(* IEC 61131-3 sources: JingjiangMoonbox/Application/Application/数据类型/通讯协议/月影/副主站通讯协议#1, 7 files *)

(* ---- StParam_Mailbox_Dep.st ---- *)
(*@CES
Name=StParam_Mailbox_Dep
Type=Gvl
TypeGuid=2db5746d-d284-4425-9f7f-2663a34b0ebc
Guid=8959721b-aa70-4a50-8488-8b5c585a49ff
HasDeclaration=True
HasImplementation=False
*)
{DECLARATION}
{attribute 'pack_mode' := '1'}
TYPE StParam_Mailbox_Dep :
STRUCT
	dwSemaphore								:DWORD;(*通讯旗语						*)

	iGirth_Uw_A								: INT; (*放A周长*)
	iGirth_Uw_B								: INT; (*放B周长*)
	iGirth_Pu								: INT;(*版周长*)
	iVelocity_Tar							: INT;(*目标速度*)
	iAI_mid_Uw								: INT;(*放料中位*)
	iAI_mid_If								: INT;(*放牵中位*)
	byDir_Uw_If_AI							: BYTE;(*放料放牵摆臂方向判断bit0:放料bit1:放牵*)
	wKp_Uw									: WORD;(*放料P*)
	wKi_Uw									: WORD;(*放料I*)
	wKd_Uw									: WORD;(*放料D*)
	wKp_If									: WORD;(*放牵P*)
	wKi_If									: WORD;(*放牵i*)
	wKd_If									: WORD;(*放牵d*)
	bySwitch_AutoCut_Uw						: BYTE;(*放料自动裁切使能开关bit0:使能；bit1:剩余卷径方式bit2:剩余米数方式*)
	iDia_PaperRoller_Uw						: INT;(*纸筒直径*10*)
	iFilmThickNess							: INT;(*料模厚度*1000*)
	wAutoMaticCutDia_Uw						: WORD;(*剩余卷径方式卷径设定*)
	wAutoMaticCutMeters_Uw					: WORD;(*剩余米数方式米数设定*)
	wActRemainFilmLenth_Uw					: WORD;(*实际剩余料长-校正纸筒直径可用*)
	iAlarm_Uw_Dia 							: INT;(*放料报警卷径设置*)
	iDelayMsec_CutterHolder					: INT;(*刀架执行时间*)
	iDelayMsec_RollerCylinder				: INT;(*压辊执行时间*)
	iDelayMsec_CutOffKnifeCylinder			: INT;(*裁刀执行时间*)
	uiMM_Roller2GummedTape					: WORD;(*压辊胶带距离*)
	uiMM_Roller2CutOfKnife					: WORD;(*压辊裁刀距离*)
	uiMM_CutOfKnife2GummedTape				: WORD;(*裁刀胶带距离*)
	iCoefCut_FilmVolPerimeter_Uw			: INT;(*放料裁切圈数*)
	iStepVariation4ChangeTime				: INT; (* 2018.9.30.100457/用来步进胶辊延时和裁刀延时的变化量 *)
	bySwitch_Compensate_Uw					: BYTE;(*放料翻转架补偿开关：Bit0:补偿开启,bit1:方向取反,bit2:0弧度确认*)
	wDiam_Tower_Uw							: WORD;(*放料翻转架的直径|mm*)
	wDiam_NextRoller_Uw						: WORD;(*放料翻转架下个辊的直径|mm*)
	wXPos_NextRoller_Uw						: WORD;(*放料翻转架下个辊的X位置|mm|翻转架中心作为坐标系0点*)
	wYPos_NextRoller_Uw						: WORD;(*放料翻转架下个辊的Y位置|mm|翻转架中心作为坐标系0点*)
	wDiam_DeflectorRoller_Uw				: WORD;(*翻料架上导向辊的直径|mm*)
	wDiam_DeflectorRollPos_Uw				: WORD;(*ABjuli翻料架的导向辊圆心运动直径|距离翻转架圆心=该值/2|mm*)
	byDiamMeasureTypeId						: BYTE;(*卷径测量方式=0：电位器=1 编码器=2 超声波(I)=3 超声波(S)=4 *)
	iStdVol_Diam_1							: INT;
	iStdVol_Diam_2							: INT;
	iStdVol_Diam_3							: INT;
	iStdVol_Diam_4							: INT;
	dwStdVol_Volt_AxisA_1					: DWORD;
	dwStdVol_Volt_AxisA_2					: DWORD;
	dwStdVol_Volt_AxisA_3					: DWORD;
	dwStdVol_Volt_AxisA_4					: DWORD;
	iStdVol_Coef_Axis_1						: INT;(* 卷径测量系数*1000 *)
	iStdVol_Coef_Axis_2						: INT;
	iStdVol_Coef_Axis_3						: INT;
	byIsDebug_DiaMeasureArea_Uw				: BYTE;
	bySwitch_DiaMeasure						: BYTE;(*bit0:自动卷径开关bit1:双轴biw2:弧面bit3:调试模式*)
	bySwitch_Enc_Uw							: BYTE;(*放料编码器标定相关bit0:双轴系数bit1:调试模式
								bit2:定位写入bit3:最小径写入*)
	(*修改变量名-放料人机屏的一些按钮通讯@2023.09.21.103603*)
	wButton_Uw 								: WORD;
	//到这里上面总共103字节||增加预留47||放牵预计总共150字节双向通讯||不够还可以扩展，总量不超过480
	abyRsv_Deputy							: ARRAY [1..47] OF BYTE;
(*以上为放牵|放料人机需要内容2025.11.16.133721||下面存放1色人机屏内容*)
	wButtonFun_Lamp_Unit					:WORD ;(*HMI界面按钮及指示灯			*)
	wSwitchFun_Unit							:WORD ;(*界面开关*)
	rStep_Pressure_Prn_Net					:REAL ;(*版辊网辊按钮步进量				*)
	rLong_Step_Roller_Pressure				:REAL ;(*色组压力控制长步进值			*)
	rShort_Step_Roller_Pressure				:REAL ;(*色组压力控制短步进值			*)
	wAirInletWindDoorValue					:WORD ;(*进风口风门开度值				*)
	wAirExhaustWindDoorValue				:WORD ;(*排风口风门开度值				*)
	wAirReturnWindDoorValue					:WORD ;(*回风口风门开度值				*)
	dwCtlBits_UnitBaseCraft					:DWORD;(*界面工艺开关及状态				*)
	wHz_UnitInkRoller_ManuallySet			:WORD ;(*递墨辊手动频率					*)
	wCoeff_UnitInkRoller_Auto				:WORD ;(*递墨辊自动系数					*)
	wHz_UnitScraper_ManuallySet				:WORD ;(*刮刀手动频率					*)
	wCoeff_UnitScraper_Auto					:WORD ;(*刮刀自动系数					*)
	wHz_UnitHotWind							:WORD ;(*热风频率						*)
	wHz_UnitHotWind_2						:WORD ;(*热风2频率						*)
	wSV_UnitTemCtl							:WORD ;(*加热设定温度					*)
	wUnit_output_I							:WORD ;(*IO监控输出1					*)
	wUnit_output_II							:WORD ;(*IO监控输出2					*)
	rHz_AxisAirBlowning_ManuallySet			: REAL;
	rHz_AxisAirExhaust_ManuallySet			: REAL;

END_STRUCT
END_TYPE

{IMPLEMENTATION}

(* ---- StPdu_Dn_91_Dep.st ---- *)
(*@CES
Name=StPdu_Dn_91_Dep
Type=Gvl
TypeGuid=2db5746d-d284-4425-9f7f-2663a34b0ebc
Guid=7bb09e6f-1753-4b92-a80e-e9a248fce2c8
HasDeclaration=True
HasImplementation=False
*)
{DECLARATION}
{attribute 'pack_mode' := '1'}
TYPE StPdu_Dn_91_Dep :
STRUCT
	byUnitId					:BYTE  ;(*机组号+系ID(最高位为系ID)*)
	rGirth_Sam					:REAL  ;(*采样版周长*)
	uiNum_Sam					:WORD  ;(*采样减速比分子*)
	uiDen_Sam					:WORD  ;(*采样减速比分母*)
	byCurrUsrLevel				:BYTE  ;(*用户权限*)
	iCompanyId					:INT   ;(*用户编号*)
	byLanguageId				:BYTE  ;(*语言选择*)
	byMinutes_ScrAutoSleep		:BYTE  ;(*屏幕休眠时间*)
	wUnit_input_I				:WORD  ;(*色组IO输入1*)
	wUnit_input_II				:WORD  ;(*色组IO输入2*)
	wUnit_input_III				:WORD  ;(*色组IO输入3*)
	wVelocity					:WORD  ;(*主机速度，单位0.1m/min*)
	wVel_Axis					:WORD  ;(*轴速度，单位0.1m/min*)
//	wComplexBit					:WORD  ;(*复合控制位描述*)
	wAxis_RollerDn				:WORD  ;(*轴压辊状态(bit0-1U,bit15-16U)*)
	wAxis_Alarm_Prn				:WORD  ;(*色组版辊报警状态(bit0-1U,bit15-16U)*)
	dwAlarmCode					:DWORD ;(*轴报警码*)
	wComplexFlag_AxisInching	:WORD  ;(*所有轴的单运行状态*)
	wComplexFlag_Linkage		:WORD  ;(*所有轴的联动状态*)
	wComplexFlag_Estop			:DWORD ;(*所有轴的急停状态*)
	wHMI_SwitchSts				:WORD  ;(*色组人机界面开关状态*)
	wSts_HorzManuPreReg			:WORD  ;(*横向手动预套准状态*)
	iPos_HorzManuPreReg			:INT   ;(*横向手动预套准位置*)
(*2025.8.6.205703增加*)
	bySts_Flag					:BYTE;(*色组状态*)
(*	dwAxis_SkipTheHeader 		:DWORD;(*让料头标志*)*)
	bySts_Machine				:BYTE;
	(*
		bit0: 印刷标志
		bit1: 空转标志
		bit2:
	*)
	//2025.11.14.155203||把误差状态发到从站，用于从站人机屏保实现9-1=8；
	byErrSts_V					: BYTE;
//用两个预留放低通滤波频率2025.11.15.132130|niu.j|8-2=6
	//Filter原本的wRsv在这里改一下改为从站精采样数据低通滤波频率
	uilowpasscutoff_hz				:UINT;

	abyRsv_91					:ARRAY [1..6] OF BYTE  ;(*预留空间*)
END_STRUCT
END_TYPE

{IMPLEMENTATION}

(* ---- StPdu_Dn_92_Dep.st ---- *)
(*@CES
Name=StPdu_Dn_92_Dep
Type=Gvl
TypeGuid=2db5746d-d284-4425-9f7f-2663a34b0ebc
Guid=436053ad-f3f5-434c-88e4-1b7334a4af27
HasDeclaration=True
HasImplementation=False
*)
{DECLARATION}
{attribute 'pack_mode' := '1'}
TYPE StPdu_Dn_92_Dep :
STRUCT
	iCurveViewMaxRange				:INT;(*误差曲线量程上限		*)
	bySignalGain					:BYTE;(*光电眼IO控制			*)
	byMarkTypeId					:BYTE;(*标记形式				*)
	byMarkArrangeModalId			:BYTE;(*标记排列形式			*)
	byFakeThreshold_V				:BYTE;(*纵向飞点阀值@丝			*)
	byFakeThreshold_H				:BYTE;(*横向飞点阀值@丝			*)
	rAlarm_V						:REAL;(*纵向报警值@mm			*)
	rAlarm_H						:REAL;(*横向报警值@mm			*)
	byAve_v_extra_V					:BYTE;(*套色误差显示平均次数	*)
	byAve_v_extra_H					:BYTE;(*套色误差显示平均次数	*)
(*	dwFlag_Sts						: DWORD;(* 状态标志 *)
(*												/bit0.纵向自动 *)
(*												/bit1.横向自动
												/bit9.双极性*)
(*												/ *)
*)
	iGateWidthPhy					: INT ;(*波门宽度				*)
	byTriangleMark_SideC			: BYTE;(*梯形标记三角形纵向边长	*)
	byTriangleMark_SideB			: BYTE;(*梯形标记三角形横向边长	*)
	bySysSamplePrecision			: BYTE;(*系统采样精度			*)
	byArcFineSampleType				: BYTE;(*套色采样方式			*)
	iSampleCfgParam_ctl				: INT ;(*采样控制参数里的ctl		*)
	byColorIdCurrent				: BYTE;(*当前色序				*)
	byColorIdFollow					: BYTE;(*跟踪色序				*)
	abyColorIdList					: ARRAY [1..16] OF BYTE;(*色序列表				*)
	//bySignalSelect					:BYTE;(*光纤电眼信号选择		*)
	xEnable_Arc						: BOOL;(*套印使能开关			*)
	uiSource_Light_T1_Cur			: UINT;
	uiSource_Light_T2_Cur			: UINT;
	abyRsv_92						: ARRAY [1..9] OF BYTE;(*套色参数预留			*)
END_STRUCT
END_TYPE

{IMPLEMENTATION}

(* ---- StPdu_Dn_93_Dep.st ---- *)
(*@CES
Name=StPdu_Dn_93_Dep
Type=Gvl
TypeGuid=2db5746d-d284-4425-9f7f-2663a34b0ebc
Guid=233641f5-af31-41e2-841e-6ff9f436d5aa
HasDeclaration=True
HasImplementation=False
*)
{DECLARATION}
{attribute 'pack_mode' := '1'}
TYPE StPdu_Dn_93_Dep :
STRUCT
	dwControlComplexBits		:DWORD;(*开关状态			*)
	wHz_UnitInkRoller_CurrWR	:WORD ;(*递墨辊最终写入频率	*)
	wHz_UnitScraper_CurrWR		:WORD ;(*刮刀写入频率		*)
	wHz_UnitHotWind_CurrWR		:WORD ;(*热风写入频率		*)
	wHz_UnitHotWind2_CurrWR		:WORD ;(*热风2写入频率		*)
	rPV_UnitTemCtl				:REAL ;(*当前温度			*)
	wSTS_UnitTemCtl				:WORD ;(*温控状态			*)
(*2025.8.6.212214增加*)
	wHotWind_Print				:WORD;(*热风打开色组号*)
	byDriverType_Hor			:BYTE;(*横向的驱动器类型*)
	wPulseCtlInf  				:WORD;(*脉冲控制信息*)
	wPulse_1r					:WORD;(*1圈的脉冲数*)
	byPulseCtl_DisPerPulse 		:BYTE;(*单位脉冲距离*)
	byPulseCtlBit 				:BYTE;(*脉冲控制位*)
	abyRsv_93					:ARRAY [1..30] OF BYTE ;(*工艺参数预留		*)
END_STRUCT
END_TYPE

{IMPLEMENTATION}

(* ---- StPdu_Dn_94_Dep.st ---- *)
(*@CES
Name=StPdu_Dn_94_Dep
Type=Gvl
TypeGuid=2db5746d-d284-4425-9f7f-2663a34b0ebc
Guid=28ccc25b-e1b3-40e8-9cb7-612afea4cc4b
HasDeclaration=True
HasImplementation=False
*)
{DECLARATION}
{attribute 'pack_mode' := '1'}
TYPE StPdu_Dn_94_Dep :
STRUCT
	rPos_M_Prn_HandWheelCtl		:REAL;(*版辊压力操作侧位置-手轮显示						*)
	rPos_G_Prn_HandWheelCtl		:REAL;(*版辊压力传动侧位置-手轮显示						*)
	rPos_M_Net_HandWheelCtl		:REAL;(*网辊压力操作侧位置-手轮显示						*)
	rPos_G_Net_HandWheelCtl		:REAL;(*网辊压力传动侧位置-手轮显示						*)
	rPos_PrnRoller_Pressure_M	:REAL;(*版辊压力操作侧实时位置							*)
	rPos_PrnRoller_Pressure_G	:REAL;(*版辊压力传动侧实时位置							*)
	rPos_NetRoller_Pressure_M	:REAL;(*网辊压力操作侧实时位置							*)
	rPos_NetRoller_Pressure_G	:REAL;(*网辊压力传动侧实时位置							*)
	byCtlId_HandWheel			:BYTE;(*手轮控制ID										*)
	byCtlSts_HandWheel			:BYTE;(*手轮控制状态									*)
	wAxis_Alarm_Net				:WORD;(*色组网辊报警状态(bit0-1U,bit15-16U)				*)
	wAxis_Alarm_Bottom			:WORD;(*色组底辊报警状态(bit0-1U,bit15-16U)				*)
	wAxis_Alarm_Prn_M			:WORD;(*色组版辊压力操作侧报警状态(bit0-1U,bit15-16U)	*)
	wAxis_Alarm_Prn_G			:WORD;(*色组版辊压力传动侧报警状态(bit0-1U,bit15-16U)	*)
	wAxis_Alarm_Net_M			:WORD;(*色组网辊压力操作侧报警状态(bit0-1U,bit15-16U)	*)
	wAxis_Alarm_Net_G			:WORD;(*色组网辊压力传动侧报警状态(bit0-1U,bit15-16U)	*)
	wAxis_Alarm_Other			:WORD;(*整机其他轴报警状态								*)
	abyRsv_93					:array [1..9] of BYTE;(*柔印参数预留									*)
END_STRUCT
END_TYPE

{IMPLEMENTATION}

(* ---- StPdu_Dn_95_Dep.st ---- *)
(*@CES
Name=StPdu_Dn_95_Dep
Type=Gvl
TypeGuid=2db5746d-d284-4425-9f7f-2663a34b0ebc
Guid=d2f57c01-a40d-42ce-9084-08d4e05e4b23
HasDeclaration=True
HasImplementation=False
*)
{DECLARATION}
{attribute 'pack_mode' := '1'}
TYPE StPdu_Dn_95_Dep :
STRUCT
END_STRUCT
END_TYPE

{IMPLEMENTATION}

(* ---- StPdu_Up_05_Dep.st ---- *)
(*@CES
Name=StPdu_Up_05_Dep
Type=Gvl
TypeGuid=2db5746d-d284-4425-9f7f-2663a34b0ebc
Guid=6633295c-2f3d-4871-ab72-dbe78eb86074
HasDeclaration=True
HasImplementation=False
*)
{DECLARATION}
{attribute 'pack_mode' := '1'}
TYPE StPdu_Up_05_Dep :
STRUCT
END_STRUCT
END_TYPE

{IMPLEMENTATION}
